Fanuc KAREL source: KT00432.KL

PROGRAM KT00432
%NOLOCKGROUP
VAR
  P1: JOINTPOS
  P2: XYZWPR
  OUT: BOOLEAN
BEGIN
    P2.Y = 2.0
  OUT = P1 > P2
END KT00432
